RoboDK station: repair_workcell.rdk

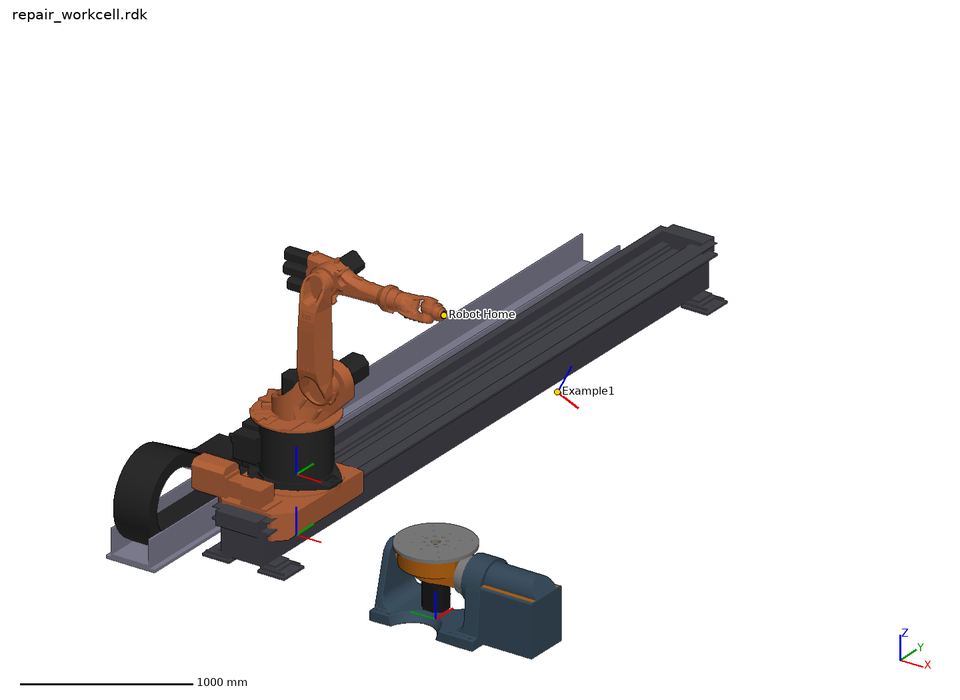
[picture v0: the station drawn from its stored meshes, robots at their saved joint values, targets as dots, program paths as lines]
Station repair_workcell (saved by RoboDK 5.5.4). Poses are relative to the parent item; angles as X-Y-Z fixed-axis rotations.
  - frame KUKA KL 250 3 Base at (0, 0, 0) mm
    - robot KUKA KL 250 3: 1 axes, payload 300 kg, reach 3600 mm, repeatability 0.02 mm
        modified DH rows (alpha deg, a mm, theta deg, d mm): -90, 0, 0, 0 linear
        joint limits [0] to [3600]; home [0]; saved at [0]
      - frame KUKA KR 6 2 Base at (0, 0, 0) mm
        - robot KUKA KR 6 2: 6 axes, payload 6 kg, reach 1611 mm, repeatability 0.05 mm, weight 235 kg
            modified DH rows (alpha deg, a mm, theta deg, d mm): 0, 0, 0, 675; -90, 260, 0, 0; 0, 680, -90, 0; -90, -35, 0, 670; 90, 0, 0, 0; -90, 0, 180, 115
            joint limits [-185, -155, -130, -350, -130, -350] to [185, 35, 154, 350, 130, 350]; home [0, -90, 90, 0, 0, 0]; saved at [0, -90, 90, -66.696, 0, 66.696]
  - frame KUKA KP2-HV500 Base at (1300, -450, 0) mm, rotated rx 0 ry 0 rz 90 deg
    - robot KUKA KP2-HV500: 2 axes
        modified DH rows (alpha deg, a mm, theta deg, d mm): 0, 0, 0, 0; -90, 0, 0, 0
        base shift (0, 0, 350) mm, rotated rx 90 ry 0 rz 0 deg
        joint limits [-135, -185] to [135, 185]; home [0, 0]; saved at [0, 0]
  - frame example at (970, 1250, 690) mm, rotated rx -25 ry 15 rz -10 deg
    - target Robot Home (joint target) at (17.79, -1550.85, 443.81) mm, rotated rx 50.97 ry 61.1 rz 57.62 deg; joints [0, -90, 90, -66.696, 0, 66.696, 0, 0, 0] of KUKA KR 6 2
    - target Example1 (joint target) at (0, 0, 0) mm; joints [-55.628, 2.21, 25.823, -252.179, 60.111, 237.174, 0, 0, 0] of KUKA KR 6 2
